(* IEC 61131-3 sources: plcassist-cli/packages/volt-lsp-iec/test-corpus/pro2193/Device/Plc Logic/Application/09 Misc/Library Manager/CmpEventMgr Implementation, 22 files *)

(* ---- EVENTCLOSE.fun ---- *)
FUNCTION EVENTCLOSE : RTS_IEC_RESULT
VAR_INPUT
	HEVENT : RTS_IEC_HANDLE;
END_VAR
VAR_IN_OUT
	RESULT : RTS_IEC_RESULT;
END_VAR
END_FUNCTION

(* ---- EVENTCLOSE2.fun ---- *)
FUNCTION EVENTCLOSE2 : RTS_IEC_RESULT
VAR_INPUT
	HEVENT : RTS_IEC_HANDLE;
END_VAR
END_FUNCTION

(* ---- EVENTCREATE.fun ---- *)
FUNCTION EVENTCREATE : RTS_IEC_HANDLE
VAR_INPUT
	EVENTID : UDINT;
	CMPIDPROVIDER : UDINT;
END_VAR
VAR_IN_OUT
	RESULT : RTS_IEC_RESULT;
END_VAR
END_FUNCTION

(* ---- EVENTCREATE2.fun ---- *)
FUNCTION EVENTCREATE2 : RTS_IEC_HANDLE
VAR_INPUT
	EVENTID : UDINT;
	CMPIDPROVIDER : UDINT;
	NCALLBACKSPOSSIBLE : UDINT;
END_VAR
VAR_IN_OUT
	RESULT : RTS_IEC_RESULT;
END_VAR
END_FUNCTION

(* ---- EVENTCREATEEVENTID.fun ---- *)
FUNCTION EVENTCREATEEVENTID : UDINT
VAR_INPUT
	EVENT : UINT;
	CLASS : UINT;
END_VAR
VAR_IN_OUT
	RESULT : RTS_IEC_RESULT;
END_VAR
END_FUNCTION

(* ---- EVENTDELETE.fun ---- *)
FUNCTION EVENTDELETE : RTS_IEC_RESULT
VAR_INPUT
	HEVENT : RTS_IEC_HANDLE;
END_VAR
VAR_IN_OUT
	RESULT : RTS_IEC_RESULT;
END_VAR
END_FUNCTION

(* ---- EVENTDELETE2.fun ---- *)
FUNCTION EVENTDELETE2 : RTS_IEC_RESULT
VAR_INPUT
	HEVENT : RTS_IEC_HANDLE;
END_VAR
END_FUNCTION

(* ---- EVENTGETCLASS.fun ---- *)
FUNCTION EVENTGETCLASS : UINT
VAR_INPUT
	EVENTID : UDINT;
END_VAR
END_FUNCTION

(* ---- EVENTGETEVENT.fun ---- *)
FUNCTION EVENTGETEVENT : UINT
VAR_INPUT
	EVENTID : UDINT;
END_VAR
END_FUNCTION

(* ---- EVENTOPEN.fun ---- *)
FUNCTION EVENTOPEN : RTS_IEC_HANDLE
VAR_INPUT
	EVENTID : UDINT;
	CMPIDPROVIDER : UDINT;
END_VAR
VAR_IN_OUT
	RESULT : RTS_IEC_RESULT;
END_VAR
END_FUNCTION

(* ---- EVENTPOST.fun ---- *)
FUNCTION EVENTPOST : RTS_IEC_RESULT
VAR_INPUT
	HEVENT : RTS_IEC_HANDLE;
	PEVENTPARAM : POINTER TO EventParam;
END_VAR
END_FUNCTION

(* ---- EVENTPOST2.fun ---- *)
FUNCTION EVENTPOST2 : RTS_IEC_RESULT
VAR_INPUT
	HEVENT : RTS_IEC_HANDLE;
	PEVENTPARAM : POINTER TO EventParam2;
END_VAR
END_FUNCTION

(* ---- EVENTPOSTBYEVENT.fun ---- *)
FUNCTION EVENTPOSTBYEVENT : RTS_IEC_RESULT
VAR_INPUT
	EVENTID : UDINT;
	CMPIDPROVIDER : UDINT;
	PEVENTPARAM : POINTER TO EventParam;
END_VAR
END_FUNCTION

(* ---- EVENTPOSTBYEVENT2.fun ---- *)
FUNCTION EVENTPOSTBYEVENT2 : RTS_IEC_RESULT
VAR_INPUT
	EVENTID : UDINT;
	CMPIDPROVIDER : UDINT;
	PEVENTPARAM : POINTER TO EventParam2;
END_VAR
END_FUNCTION

(* ---- EVENTREGISTERCALLBACK.fun ---- *)
FUNCTION EVENTREGISTERCALLBACK : RTS_IEC_HANDLE
VAR_INPUT
	HEVENT : RTS_IEC_HANDLE;
	PICALLBACK : ICmpEventCallback;
END_VAR
VAR_IN_OUT
	RESULT : RTS_IEC_RESULT;
END_VAR
END_FUNCTION

(* ---- EVENTREGISTERCALLBACK2.fun ---- *)
FUNCTION EVENTREGISTERCALLBACK2 : RTS_IEC_HANDLE
VAR_INPUT
	HEVENT : RTS_IEC_HANDLE;
	PICALLBACK : ICmpEventCallback;
	PUSERPARAMETER : POINTER TO BYTE;
END_VAR
VAR_IN_OUT
	RESULT : RTS_IEC_RESULT;
END_VAR
END_FUNCTION

(* ---- EVENTREGISTERCALLBACKFUNCTION.fun ---- *)
FUNCTION EVENTREGISTERCALLBACKFUNCTION : RTS_IEC_RESULT
VAR_INPUT
	HEVENT : RTS_IEC_HANDLE;
	PFCALLBACKFUNCTION : POINTER TO BYTE;
END_VAR
END_FUNCTION

(* ---- EVENTREGISTERCALLBACKFUNCTION2.fun ---- *)
FUNCTION EVENTREGISTERCALLBACKFUNCTION2 : RTS_IEC_RESULT
VAR_INPUT
	HEVENT : RTS_IEC_HANDLE;
	PFCALLBACKFUNCTION : POINTER TO BYTE;
	PUSERPARAMETER : POINTER TO BYTE;
END_VAR
END_FUNCTION

(* ---- EVENTREGISTEREDCALLBACKS.fun ---- *)
FUNCTION EVENTREGISTEREDCALLBACKS : UDINT
VAR_INPUT
	HEVENT : RTS_IEC_HANDLE;
END_VAR
VAR_IN_OUT
	RESULT : RTS_IEC_RESULT;
END_VAR
END_FUNCTION

(* ---- EVENTUNREGISTERCALLBACK.fun ---- *)
FUNCTION EVENTUNREGISTERCALLBACK : RTS_IEC_RESULT
VAR_INPUT
	HEVENT : RTS_IEC_HANDLE;
	HINTERFACE : RTS_IEC_HANDLE;
END_VAR
END_FUNCTION

(* ---- EVENTUNREGISTERCALLBACKFUNCTION.fun ---- *)
FUNCTION EVENTUNREGISTERCALLBACKFUNCTION : RTS_IEC_RESULT
VAR_INPUT
	HEVENT : RTS_IEC_HANDLE;
	PFCALLBACKFUNCTION : POINTER TO BYTE;
END_VAR
END_FUNCTION

(* ---- EVENTUNREGISTERCALLBACKFUNCTION2.fun ---- *)
FUNCTION EVENTUNREGISTERCALLBACKFUNCTION2 : RTS_IEC_RESULT
VAR_INPUT
	HEVENT : RTS_IEC_HANDLE;
	PFCALLBACKFUNCTION : POINTER TO BYTE;
	PUSERPARAMETER : POINTER TO BYTE;
END_VAR
END_FUNCTION
